Fanuc KAREL source: KA00038.KL

PROGRAM KA00038
%NOLOCKGROUP
VAR
  SRC: STRING[80]
  DST: REAL
BEGIN
  SRC = 'A'
  DST = SRC
END KA00038
